{attribute 'qualified_only'}
VAR_GLOBAL
    stInputs  : ST_MachineInputs;
    stOutputs : ST_MachineOutputs;
    stCommand : ST_MachineCommand;
    stStatus  : ST_MachineStatus;
    stStationEvents   : ARRAY[0..4] OF ST_StationEvents;
    stEventsAssigment : ST_EventsAssigmentGeneral;
    astActiveEvents   : ARRAY[0..50] OF ST_ActiveEvents;
    sSystemTime       : STRING(255);
    sSystemDate       : STRING(255);
    bMachineFault     : BOOL;
    bCycleStopRequest : BOOL;
    // Manual index warnings: presentation only, never Fault/Stop requests.
    bManualIndexBlockVision : BOOL;
    bManualIndexBlockHeat : BOOL;
    bManualIndexBlockPatch : BOOL;
    bManualIndexBlockOther : BOOL;
    sManualIndexVisionReason : STRING(160);
    sManualIndexOtherReason : STRING(160);
    bManualCameraRecoveryFailed : BOOL;
    bVisionManualCameraWarning : BOOL;
    bVisionManualGridWarning : BOOL;
    bVisionManualGridActive : BOOL;
END_VAR
VAR_GLOBAL CONSTANT
    // Per-nest Heat Stake product-quality warning identity (not a machine fault).
    udiHeatStakePatchMissingAlertCode : UDINT := 1201;
END_VAR

(* stored: Version 1.1.0.1, ProductVersion 3.1.4026.18
   GVL GVL_MASTER: Id {9970f182-028c-4164-bcf7-ddc50b57d0ed} *)
